(* IEC 61131-3 sources: Elmo_Master/Lasal_PRG/Elmo_EtherCAT_Test_4Axis/Class/_TCPIPServer (part 2) *)

        (*================================================================*)
        SVR_TCP_CMD_CLOSESOCKETTYPE:
        (*================================================================*)
          case SubCmd of
            (*==================================================*)
            SVR_TCP_CLOSESOCKETTYPE:
            (*==================================================*)
              pConn^.CloseSocketType := ParaValue$UDINT;
            (*==================================================*)
            else // - INVALID SUB COMMAND
            (*==================================================*)
              Retcode := TCP_SVR_ERR_SET_PARA_INVALID_SUB_CMD;
          end_case;

        (*================================================================*)
        else // - INVALID COMMAND
        (*================================================================*)
          Retcode := TCP_SVR_ERR_SET_PARA_INVALID_CMD;

      end_case;
    else
      Retcode := TCP_SVR_ERR_INVALID_SOCKET;
    end_if;
  else
    Retcode := TCP_SVR_ERR_INVALID_SOCKET;
  end_if;

END_FUNCTION

FUNCTION VIRTUAL GLOBAL _TCPIPServer::ReadMainParameter
	VAR_INPUT
		Cmd 	: DINT;
		SubCmd 	: DINT;
		pParaValue 	: ^DINT;
	END_VAR
	VAR_OUTPUT
		Retcode 	: DINT;
	END_VAR

  Retcode := TCP_SVR_NO_ERROR;

  if (usInit > 0) then
    case Cmd of
      (*================================================================*)
      SVR_TCP_CMD_SETSOCKOPT:
      (*================================================================*)
        case SubCmd of
          (*==================================================*)
          SVR_TCP_SOCKOPT_NAGLE:
          (*==================================================*)
            if (MainSockOpt.Nagle = false) then
              pParaValue^ := 0;
            else
              pParaValue^ := 1;
            end_if;
          (*==================================================*)
          SVR_TCP_SOCKOPT_KEEPALIVE:
          (*==================================================*)
            if (MainSockOpt.KeepAlive = false) then
              pParaValue^ := 0;
            else
              pParaValue^ := 1;
            end_if;
          (*==================================================*)
          SVR_TCP_SOCKOPT_DELAYEDACK:
          (*==================================================*)
            if (MainSockOpt.DelayedAck = false) then
              pParaValue^ := 0;
            else
              pParaValue^ := 1;
            end_if;
          (*==================================================*)
          SVR_TCP_SOCKOPT_REUSEADDR:
          (*==================================================*)
            if (MainSockOpt.ReuseAddr = false) then
              pParaValue^ := 0;
            else
              pParaValue^ := 1;
            end_if;
          (*==================================================*)
          else // - INVALID SUB COMMAND
          (*==================================================*)
            Retcode := TCP_SVR_ERR_SET_PARA_INVALID_SUB_CMD;
        end_case;

      (*================================================================*)
      SVR_TCP_CMD_TASKPRIO:
      (*================================================================*)
        case SubCmd of
          (*==================================================*)
          SVR_TCP_SUB_CMD_TASKPRIO:
          (*==================================================*)
            pParaValue^ := AP_TaskPriority$DINT;
          (*==================================================*)
          else // - INVALID SUB COMMAND
          (*==================================================*)
            Retcode := TCP_SVR_ERR_SET_PARA_INVALID_SUB_CMD;
        end_case;

      (*================================================================*)
      SVR_TCP_CMD_KEEPALIVEPARA: // - ASYNC TASK PRIORITY
      (*================================================================*)
        case SubCmd of
          (*==================================================*)
          SVR_TCP_KEEPALIVE_KEEPIDLE:
          (*==================================================*)
            pParaValue^ := KeepAlivePara.keepIDLE;
          (*==================================================*)
          SVR_TCP_KEEPALIVE_KEEPINTVL:
          (*==================================================*)
            pParaValue^ := KeepAlivePara.keepINTVL;
          (*==================================================*)
          SVR_TCP_KEEPALIVE_KEEPCNT:
          (*==================================================*)
            pParaValue^ := KeepAlivePara.keepCNT;
          (*==================================================*)
          else // - INVALID SUB COMMAND
          (*==================================================*)
            Retcode := TCP_SVR_ERR_SET_PARA_INVALID_SUB_CMD;
        end_case;

      (*================================================================*)
      SVR_TCP_CMD_CLOSESOCKETTYPE:
      (*================================================================*)
        case SubCmd of
          (*==================================================*)
          SVR_TCP_CLOSESOCKETTYPE:
          (*==================================================*)
            pParaValue^$UDINT := CloseSocketType;
          (*==================================================*)
          else // - INVALID SUB COMMAND
          (*==================================================*)
            Retcode := TCP_SVR_ERR_SET_PARA_INVALID_SUB_CMD;
        end_case;

      (*================================================================*)
      else // - INVALID COMMAND
      (*================================================================*)
        Retcode := TCP_SVR_ERR_SET_PARA_INVALID_CMD;

    end_case;
  else
    Retcode := TCP_SVR_ERR_MAIN_INIT;
  end_if;

END_FUNCTION

FUNCTION VIRTUAL GLOBAL _TCPIPServer::ReadSocketParameter
	VAR_INPUT
		dSock 	: DINT;
		Cmd 	: DINT;
		SubCmd 	: DINT;
		pParaValue 	: ^DINT;
	END_VAR
	VAR_OUTPUT
		Retcode 	: DINT;
	END_VAR
VAR
	pConn       : ^_CONNECTION;
END_VAR

  Retcode := TCP_SVR_NO_ERROR;

  if (CheckSocketValid(dSock, (#pConn)$^pVoid) = true) then
    if (pConn <> NIL) then
      case Cmd of
        (*================================================================*)
        SVR_TCP_CMD_SETSOCKOPT:
        (*================================================================*)
          case SubCmd of
            (*==================================================*)
            SVR_TCP_SOCKOPT_NAGLE:
            (*==================================================*)
              if (pConn^.ConnSockOpt.Nagle = false) then
                pParaValue^ := 0;
              else
                pParaValue^ := 1;
              end_if;
            (*==================================================*)
            SVR_TCP_SOCKOPT_KEEPALIVE:
            (*==================================================*)
              if (pConn^.ConnSockOpt.KeepAlive = false) then
                pParaValue^ := 0;
              else
                pParaValue^ := 1;
              end_if;
            (*==================================================*)
            SVR_TCP_SOCKOPT_DELAYEDACK:
            (*==================================================*)
              if (pConn^.ConnSockOpt.DelayedAck = false) then
                pParaValue^ := 0;
              else
                pParaValue^ := 1;
              end_if;
            (*==================================================*)
            SVR_TCP_SOCKOPT_REUSEADDR:
            (*==================================================*)
              if (pConn^.ConnSockOpt.ReuseAddr = false) then
                pParaValue^ := 0;
              else
                pParaValue^ := 1;
              end_if;
            (*==================================================*)
            else // - INVALID SUB COMMAND
            (*==================================================*)
              Retcode := TCP_SVR_ERR_SET_PARA_INVALID_SUB_CMD;
          end_case;

        (*================================================================*)
        SVR_TCP_CMD_KEEPALIVEPARA: // - ASYNC TASK PRIORITY
        (*================================================================*)
          case SubCmd of
            (*==================================================*)
            SVR_TCP_KEEPALIVE_KEEPIDLE:
            (*==================================================*)
              pParaValue^ := pConn^.KeepAlivePara.keepIDLE;
            (*==================================================*)
            SVR_TCP_KEEPALIVE_KEEPINTVL:
            (*==================================================*)
              pParaValue^ := pConn^.KeepAlivePara.keepINTVL;
            (*==================================================*)
            SVR_TCP_KEEPALIVE_KEEPCNT:
            (*==================================================*)
              pParaValue^ := pConn^.KeepAlivePara.keepCNT;
            (*==================================================*)
            else // - INVALID SUB COMMAND
            (*==================================================*)
              Retcode := TCP_SVR_ERR_SET_PARA_INVALID_SUB_CMD;
          end_case;

        (*================================================================*)
        SVR_TCP_CMD_CLOSESOCKETTYPE:
        (*================================================================*)
          case SubCmd of
            (*==================================================*)
            SVR_TCP_CLOSESOCKETTYPE:
            (*==================================================*)
              pParaValue^$UDINT := pConn^.CloseSocketType;
            (*==================================================*)
            else // - INVALID SUB COMMAND
            (*==================================================*)
              Retcode := TCP_SVR_ERR_SET_PARA_INVALID_SUB_CMD;
          end_case;

        (*================================================================*)
        else // - INVALID COMMAND
        (*================================================================*)
          Retcode := TCP_SVR_ERR_SET_PARA_INVALID_CMD;

      end_case;
    else
      Retcode := TCP_SVR_ERR_INVALID_SOCKET;
    end_if;
  else
    Retcode := TCP_SVR_ERR_INVALID_SOCKET;
  end_if;

END_FUNCTION

FUNCTION _TCPIPServer::CheckSocketValid
	VAR_INPUT
		dSock 	: DINT;
		ppConn 	: ^pVoid;
	END_VAR
	VAR_OUTPUT
		Retcode 	: BOOL;
	END_VAR
VAR
	i         : USINT;
END_VAR

  Retcode := false;
  if (ppConn <> NIL) then
    ppConn^ := NIL;
  end_if;

  for i := 0 to (MaxConn-1) do
    if (SocketArray[i].dSocket = dSock) then
      if (ppConn <> NIL) then
        ppConn^ := (#SocketArray[i])$^void;
      end_if;
      Retcode := true;
      exit;
    end_if;
  end_for;

END_FUNCTION

FUNCTION GLOBAL _TCPIPServer::AddInterface
	VAR_INPUT
		thispointer 	: ^void;
	END_VAR
	VAR_OUTPUT
		dRetcode 	: DINT;
	END_VAR

  // check pointer
  if thispointer <> NIL then
    // only one Interface allowed
    if pThisInterface = NIL then
      // save thispointer for callbacks.
      pThisInterface := thispointer$^_TCPIPServerInterface;
      dRetcode := 1;
      bdStatus.ErrorNoUserInterface := FALSE;
    else
      // there is already on interface connected
      dRetcode := -1;
    end_if;
  else
    // invalid Pointer
    dRetcode := -2;
  end_if;

END_FUNCTION
